(* Cycle Running Blinky *)

PROGRAM main
  VAR
    RunState AT %MX0.0 : BOOL; (* Input Variable *)
    CycleOn AT %QX0.2 : BOOL;
    TON0 : TON;
    TOF0 : TOF;
  END_VAR

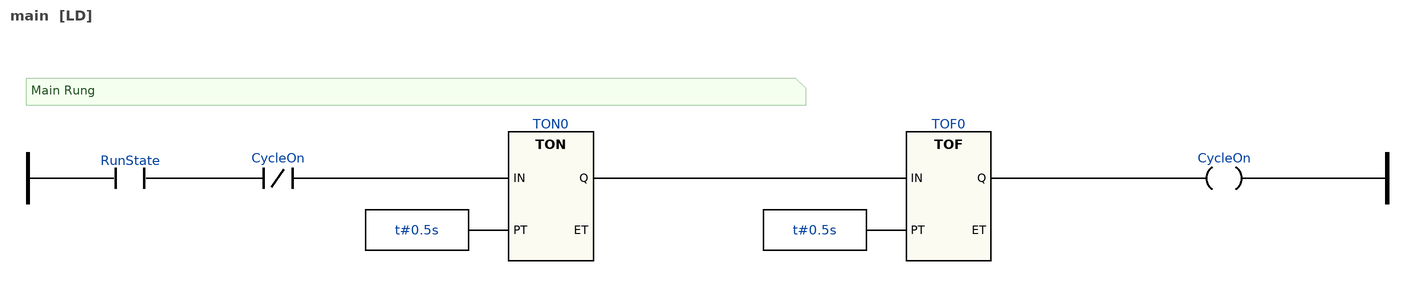
(* LD diagram, written out as Structured Text *)
(* Main Rung *)
TON0(IN := RunState AND NOT CycleOn, PT := t#0.5s);
TOF0(IN := TON0.Q, PT := t#0.5s);
CycleOn := TOF0.Q;
END_PROGRAM
